(* IEC 61131-3 sources: IRIS-Project/LASAL CONTROL SOFTWARE/LasalProject_2025_09_12/Network/Comunicazione_ModBus, 1 file *)

(* ---- ONE_Comunicazione_ModBus_Table.st ---- *)
#define OBJECTS_CONFIG

//Define part of class _TCPIP_SERVER
#ifndef OS_VERSION_MIN_SALAMANDER
    #define OS_VERSION_MIN_SALAMANDER          0x9000
  #endif
  #define TCP_SVR_NO_ERROR                          0

  #define TCP_SVR_ERR_INVALID_SOCKET            -1

  #define TCP_SVR_ERR_SET_PARA_INVALID_CMD     -10
  #define TCP_SVR_ERR_SET_PARA_INVALID_SUB_CMD -11

  #define TCP_SVR_ERR_TASK_ALREADY_EXIST       -12

  // - RETURN VALUES PRIVATE METHOD Read_AP_TaskPeriod
  #define TCP_SVR_ERR_TASK_TIME_NO_APP            -31
  #define TCP_SVR_ERR_TASK_TIME_WRONG_TASK_TYPE   -33
  #define TCP_SVR_ERR_TASK_TIME_OBJ_NOT_FOUND     -35

  // - RETURN VALUES PRIVATE METHOD Read_LSLOBJ_CRC32
  #define TCP_SVR_ERR_GET_LSLOBJ_NAME             -20
  #define TCP_SVR_ERR_INVALID_POINTER             -21

  // - RETURN VALUES PRIVATE METHOD AP_TaskCreate
  #define TCP_SVR_ERR_TASK_CREATE                 -40

  // - RETURN VALUES PRIVATE METHOD AP_SemaCreate
  #define TCP_SVR_ERR_SEMA_CREATE                 -50
  #define TCP_SVR_ERR_SEMA_INVALID_IDX            -51
  #define TCP_SVR_ERR_SEMA_INVALID_NAME           -52

  #define TCP_SVR_SEND_BUFFER_EMPTY               -6
  #define TCP_SVR_ERR_SEND_BUFFER_FATAL_ERROR     -7

  #define TCP_SVR_SEND_BUFFER_FULL      -4

  #define TCP_SVR_SOCK_INFO_CONNECT                 1
  #define TCP_SVR_SOCK_INFO_DISCONNECT              0

  #define TCP_SVR_ERR_GROUP_OS                      0
  #define TCP_SVR_ERR_GROUP_AP                      1

  #define TCP_SVR_ERR_CODE_AP_TIMEOUT              -1

  #ifndef INIT_FIRSTSCAN
    #define INIT_FIRSTSCAN                         12
  #endif

  #ifndef AP_TASK_PRIORITY_DEFAULT
    #define AP_TASK_PRIORITY_DEFAULT               14
  #endif

  #define TCP_SVR_ERR_MAIN_INIT                   -90

  #define TCP_SVR_ERR_MAX_CONN                    -80

  #ifndef KEEPALIVE_INTERVAL_DEFAULT
    #define KEEPALIVE_INTERVAL_DEFAULT           7200
  #endif

  #ifndef KEEPALIVE_RETRYTIME_DEFAULT
    #define KEEPALIVE_RETRYTIME_DEFAULT            75
  #endif

  #ifndef KEEPALIVE_RETRYCNT_DEFUALT
    #define KEEPALIVE_RETRYCNT_DEFUALT             10
  #endif

  #ifndef CLOSE_SOCKET_TYPE_DEFAULT
    #define CLOSE_SOCKET_TYPE_DEFAULT               0
  #endif
#include "..\..\Class\_TCPIP_SERVER\SalamanderDelay.h"
#include "..\..\Source\MB_Definitions.h"
#include "..\..\Runtime\%LASALAPPDATA%\Runtime\Include\LSL\lsl_st_mt.h"

FUNCTION GLOBAL TAB ONE_Comunicazione_ModBus
-1$UINT, 0$UINT,
0$UINT, 0$UINT,

15$UDINT,
TO_UDINT(916194998), "_CheckSum", 1$UINT, 0$UINT, 3$UINT,
TO_UDINT(1436589033), "_ModBusTCPSLAVE", 1$UINT, 36$UINT, 3$UINT,
TO_UDINT(26234884), "_TCPIP_SERVER", 1$UINT, 38$UINT, 0$UINT,
TO_UDINT(2897291062), "ASCII_BIN", 1$UINT, 21$UINT, 3$UINT,
TO_UDINT(1067997253), "ControlloServerModBus", 0$UINT, 0$UINT, 3$UINT,
TO_UDINT(3132304963), "HoldingRegister", 0$UINT, 0$UINT, 1$UINT,
TO_UDINT(3014633822), "HoldingRegister_2", 0$UINT, 0$UINT, 1$UINT,
TO_UDINT(3299383752), "HoldingRegister_3", 0$UINT, 0$UINT, 1$UINT,
TO_UDINT(418069068), "InputRegister", 0$UINT, 0$UINT, 3$UINT,
TO_UDINT(2225119864), "MerkerEx", 1$UINT, 22$UINT, 9$UINT,
TO_UDINT(3487210139), "MPS", 0$UINT, 0$UINT, 1$UINT,
TO_UDINT(4105514139), "Rack12V", 0$UINT, 0$UINT, 1$UINT,
TO_UDINT(1850111279), "String", 1$UINT, 11$UINT, 9$UINT,
TO_UDINT(2898603620), "StringInternal", 1$UINT, 85$UINT, 0$UINT,
TO_UDINT(3232495061), "VirtualBaseInit", 1$UINT, 3$UINT, 0$UINT,

1$UINT, TO_UDINT(966565638), "_MODBUSTCPSLAVE1\_BASE\CHECKSUM",
1$UINT, TO_UDINT(273951732), "_MODBUSTCPSLAVE2\_BASE\CHECKSUM",
1$UINT, TO_UDINT(3191650917), "_MODBUSTCPSLAVE3\_BASE\CHECKSUM",

_NO_ATTR, TO_UDINT(1516180976), "_MODBUSTCPSLAVE1",
_NO_ATTR, TO_UDINT(3277210698), "_MODBUSTCPSLAVE2",
_NO_ATTR, TO_UDINT(3025237212), "_MODBUSTCPSLAVE3",

_NO_ATTR, TO_UDINT(3586366131), "ASCII_BIN2",
_NO_ATTR, TO_UDINT(2730797605), "ASCII_BIN3",
_NO_ATTR, TO_UDINT(1017134982), "ASCII_BIN4",

_NO_ATTR, TO_UDINT(2237002480), "CONTROLLOSERVERMODBUS1",
_NO_ATTR, TO_UDINT(475833162), "CONTROLLOSERVERMODBUS2",
_NO_ATTR, TO_UDINT(1801163740), "CONTROLLOSERVERMODBUS3",

_NO_ATTR, TO_UDINT(1823689907), "HOLDINGREGISTER1",

_NO_ATTR, TO_UDINT(263994605), "HOLDINGREGISTER_21",

_NO_ATTR, TO_UDINT(380046764), "HOLDINGREGISTER_31",

_NO_ATTR, TO_UDINT(4239264054), "INPUTREGISTER1",
_NO_ATTR, TO_UDINT(1705465996), "INPUTREGISTER2",
_NO_ATTR, TO_UDINT(312502298), "INPUTREGISTER3",

1$UINT, TO_UDINT(392675759), "_MODBUSTCPSLAVE1\_BASE\STRSEMANAME01\MERKEREX0",
1$UINT, TO_UDINT(2391123886), "_MODBUSTCPSLAVE1\_BASE\STRSEMANAME02\MERKEREX0",
1$UINT, TO_UDINT(2044784268), "_MODBUSTCPSLAVE1\_BASE\STRTASKNAME\MERKEREX0",
1$UINT, TO_UDINT(72349916), "_MODBUSTCPSLAVE2\_BASE\STRSEMANAME01\MERKEREX0",
1$UINT, TO_UDINT(2645401309), "_MODBUSTCPSLAVE2\_BASE\STRSEMANAME02\MERKEREX0",
1$UINT, TO_UDINT(3706226144), "_MODBUSTCPSLAVE2\_BASE\STRTASKNAME\MERKEREX0",
1$UINT, TO_UDINT(178786317), "_MODBUSTCPSLAVE3\_BASE\STRSEMANAME01\MERKEREX0",
1$UINT, TO_UDINT(2471130636), "_MODBUSTCPSLAVE3\_BASE\STRSEMANAME02\MERKEREX0",
1$UINT, TO_UDINT(3220135108), "_MODBUSTCPSLAVE3\_BASE\STRTASKNAME\MERKEREX0",

_NO_ATTR, TO_UDINT(3838738401), "MPS1",

_NO_ATTR, TO_UDINT(3841265751), "RACK12V1",

1$UINT, TO_UDINT(191419237), "_MODBUSTCPSLAVE1\_BASE\STRSEMANAME01",
1$UINT, TO_UDINT(2455864031), "_MODBUSTCPSLAVE1\_BASE\STRSEMANAME02",
1$UINT, TO_UDINT(2184963303), "_MODBUSTCPSLAVE1\_BASE\STRTASKNAME",
1$UINT, TO_UDINT(1886802310), "_MODBUSTCPSLAVE2\_BASE\STRSEMANAME01",
1$UINT, TO_UDINT(3917414460), "_MODBUSTCPSLAVE2\_BASE\STRSEMANAME02",
1$UINT, TO_UDINT(560816718), "_MODBUSTCPSLAVE2\_BASE\STRTASKNAME",
1$UINT, TO_UDINT(4021080600), "_MODBUSTCPSLAVE3\_BASE\STRSEMANAME01",
1$UINT, TO_UDINT(1990558626), "_MODBUSTCPSLAVE3\_BASE\STRSEMANAME02",
1$UINT, TO_UDINT(4136624662), "_MODBUSTCPSLAVE3\_BASE\STRTASKNAME",

//Internal connections
0$UDINT,
21$UDINT,
TO_UDINT(3), "CheckSum", TO_UDINT(0),
TO_UDINT(3), "StrTaskName", TO_UDINT(31),
TO_UDINT(3), "StrSemaName01", TO_UDINT(29),
TO_UDINT(3), "StrSemaName02", TO_UDINT(30),
TO_UDINT(4), "CheckSum", TO_UDINT(1),
TO_UDINT(4), "StrTaskName", TO_UDINT(34),
TO_UDINT(4), "StrSemaName01", TO_UDINT(32),
TO_UDINT(4), "StrSemaName02", TO_UDINT(33),
TO_UDINT(5), "CheckSum", TO_UDINT(2),
TO_UDINT(5), "StrTaskName", TO_UDINT(37),
TO_UDINT(5), "StrSemaName01", TO_UDINT(35),
TO_UDINT(5), "StrSemaName02", TO_UDINT(36),
TO_UDINT(29), "MerkerEx0", TO_UDINT(18),
TO_UDINT(30), "MerkerEx0", TO_UDINT(19),
TO_UDINT(31), "MerkerEx0", TO_UDINT(20),
TO_UDINT(32), "MerkerEx0", TO_UDINT(21),
TO_UDINT(33), "MerkerEx0", TO_UDINT(22),
TO_UDINT(34), "MerkerEx0", TO_UDINT(23),
TO_UDINT(35), "MerkerEx0", TO_UDINT(24),
TO_UDINT(36), "MerkerEx0", TO_UDINT(25),
TO_UDINT(37), "MerkerEx0", TO_UDINT(26),
0$UDINT,
21$UDINT,
TO_UDINT(3), "cTable", TO_UDINT(12), "ClassSvr",
TO_UDINT(3), "cTableInputReg", TO_UDINT(15), "ClassSvr",
TO_UDINT(3), "to_AsciiBin", TO_UDINT(6), "Obj_channel",
TO_UDINT(4), "cTable", TO_UDINT(13), "ClassSvr",
TO_UDINT(4), "cTableInputReg", TO_UDINT(16), "ClassSvr",
TO_UDINT(4), "to_AsciiBin", TO_UDINT(7), "Obj_channel",
TO_UDINT(5), "cTable", TO_UDINT(14), "ClassSvr",
TO_UDINT(5), "cTableInputReg", TO_UDINT(17), "ClassSvr",
TO_UDINT(5), "to_AsciiBin", TO_UDINT(8), "Obj_channel",
TO_UDINT(9), "oc_ModBusTCPSlave", TO_UDINT(3), "sControl",
TO_UDINT(10), "oc_ModBusTCPSlave", TO_UDINT(4), "sControl",
TO_UDINT(11), "oc_ModBusTCPSlave", TO_UDINT(5), "sControl",
TO_UDINT(29), "DataBuffer", TO_UDINT(18), "m_udLength",
TO_UDINT(30), "DataBuffer", TO_UDINT(19), "m_udLength",
TO_UDINT(31), "DataBuffer", TO_UDINT(20), "m_udLength",
TO_UDINT(32), "DataBuffer", TO_UDINT(21), "m_udLength",
TO_UDINT(33), "DataBuffer", TO_UDINT(22), "m_udLength",
TO_UDINT(34), "DataBuffer", TO_UDINT(23), "m_udLength",
TO_UDINT(35), "DataBuffer", TO_UDINT(24), "m_udLength",
TO_UDINT(36), "DataBuffer", TO_UDINT(25), "m_udLength",
TO_UDINT(37), "DataBuffer", TO_UDINT(26), "m_udLength",

//Initialization values
0$UDINT,
39$UDINT,
TO_UDINT(3), "sDisable", TO_UDINT(0),//|Comunicazione_ModBus._ModBusTCPSLAVE1.sDisable;
TO_UDINT(3), "cPort", TO_UDINT(502),//|Comunicazione_ModBus._ModBusTCPSLAVE1.cPort;
TO_UDINT(3), "cMaxConnections", TO_UDINT(0),//|Comunicazione_ModBus._ModBusTCPSLAVE1.cMaxConnections;
TO_UDINT(3), "cBufSize", TO_UDINT(100),//|Comunicazione_ModBus._ModBusTCPSLAVE1.cBufSize;
TO_UDINT(3), "cBufSizeInputReg", TO_UDINT(100),//|Comunicazione_ModBus._ModBusTCPSLAVE1.cBufSizeInputReg;
TO_UDINT(3), "cFileOrTable", TO_UDINT(2#11),//|Comunicazione_ModBus._ModBusTCPSLAVE1.cFileOrTable;
TO_UDINT(3), "cTurnBytes", TO_UDINT(1),//|Comunicazione_ModBus._ModBusTCPSLAVE1.cTurnBytes;
TO_UDINT(4), "sDisable", TO_UDINT(0),//|Comunicazione_ModBus._ModBusTCPSLAVE2.sDisable;
TO_UDINT(4), "cPort", TO_UDINT(503),//|Comunicazione_ModBus._ModBusTCPSLAVE2.cPort;
TO_UDINT(4), "cMaxConnections", TO_UDINT(0),//|Comunicazione_ModBus._ModBusTCPSLAVE2.cMaxConnections;
TO_UDINT(4), "cBufSize", TO_UDINT(100),//|Comunicazione_ModBus._ModBusTCPSLAVE2.cBufSize;
TO_UDINT(4), "cBufSizeInputReg", TO_UDINT(100),//|Comunicazione_ModBus._ModBusTCPSLAVE2.cBufSizeInputReg;
TO_UDINT(4), "cFileOrTable", TO_UDINT(2#11),//|Comunicazione_ModBus._ModBusTCPSLAVE2.cFileOrTable;
TO_UDINT(4), "cTurnBytes", TO_UDINT(1),//|Comunicazione_ModBus._ModBusTCPSLAVE2.cTurnBytes;
TO_UDINT(5), "sDisable", TO_UDINT(0),//|Comunicazione_ModBus._ModBusTCPSLAVE3.sDisable;
TO_UDINT(5), "cPort", TO_UDINT(504),//|Comunicazione_ModBus._ModBusTCPSLAVE3.cPort;
TO_UDINT(5), "cMaxConnections", TO_UDINT(0),//|Comunicazione_ModBus._ModBusTCPSLAVE3.cMaxConnections;
TO_UDINT(5), "cBufSize", TO_UDINT(100),//|Comunicazione_ModBus._ModBusTCPSLAVE3.cBufSize;
TO_UDINT(5), "cBufSizeInputReg", TO_UDINT(100),//|Comunicazione_ModBus._ModBusTCPSLAVE3.cBufSizeInputReg;
TO_UDINT(5), "cFileOrTable", TO_UDINT(2#11),//|Comunicazione_ModBus._ModBusTCPSLAVE3.cFileOrTable;
TO_UDINT(5), "cTurnBytes", TO_UDINT(1),//|Comunicazione_ModBus._ModBusTCPSLAVE3.cTurnBytes;
TO_UDINT(18), "ThreadSafe", TO_UDINT(0),//|Comunicazione_ModBus.StrSemaName01\_base\_ModBusTCPSLAVE1\MerkerEx0.ThreadSafe;
TO_UDINT(19), "ThreadSafe", TO_UDINT(0),//|Comunicazione_ModBus.StrSemaName02\_base\_ModBusTCPSLAVE1\MerkerEx0.ThreadSafe;
TO_UDINT(20), "ThreadSafe", TO_UDINT(0),//|Comunicazione_ModBus.StrTaskName\_base\_ModBusTCPSLAVE1\MerkerEx0.ThreadSafe;
TO_UDINT(21), "ThreadSafe", TO_UDINT(0),//|Comunicazione_ModBus.StrSemaName01\_base\_ModBusTCPSLAVE2\MerkerEx0.ThreadSafe;
TO_UDINT(22), "ThreadSafe", TO_UDINT(0),//|Comunicazione_ModBus.StrSemaName02\_base\_ModBusTCPSLAVE2\MerkerEx0.ThreadSafe;
TO_UDINT(23), "ThreadSafe", TO_UDINT(0),//|Comunicazione_ModBus.StrTaskName\_base\_ModBusTCPSLAVE2\MerkerEx0.ThreadSafe;
TO_UDINT(24), "ThreadSafe", TO_UDINT(0),//|Comunicazione_ModBus.StrSemaName01\_base\_ModBusTCPSLAVE3\MerkerEx0.ThreadSafe;
TO_UDINT(25), "ThreadSafe", TO_UDINT(0),//|Comunicazione_ModBus.StrSemaName02\_base\_ModBusTCPSLAVE3\MerkerEx0.ThreadSafe;
TO_UDINT(26), "ThreadSafe", TO_UDINT(0),//|Comunicazione_ModBus.StrTaskName\_base\_ModBusTCPSLAVE3\MerkerEx0.ThreadSafe;
TO_UDINT(29), "SingleRealloc", TO_UDINT(1),//|Comunicazione_ModBus._base\_ModBusTCPSLAVE1\StrSemaName01.SingleRealloc;
TO_UDINT(30), "SingleRealloc", TO_UDINT(1),//|Comunicazione_ModBus._base\_ModBusTCPSLAVE1\StrSemaName02.SingleRealloc;
TO_UDINT(31), "SingleRealloc", TO_UDINT(1),//|Comunicazione_ModBus._base\_ModBusTCPSLAVE1\StrTaskName.SingleRealloc;
TO_UDINT(32), "SingleRealloc", TO_UDINT(1),//|Comunicazione_ModBus._base\_ModBusTCPSLAVE2\StrSemaName01.SingleRealloc;
TO_UDINT(33), "SingleRealloc", TO_UDINT(1),//|Comunicazione_ModBus._base\_ModBusTCPSLAVE2\StrSemaName02.SingleRealloc;
TO_UDINT(34), "SingleRealloc", TO_UDINT(1),//|Comunicazione_ModBus._base\_ModBusTCPSLAVE2\StrTaskName.SingleRealloc;
TO_UDINT(35), "SingleRealloc", TO_UDINT(1),//|Comunicazione_ModBus._base\_ModBusTCPSLAVE3\StrSemaName01.SingleRealloc;
TO_UDINT(36), "SingleRealloc", TO_UDINT(1),//|Comunicazione_ModBus._base\_ModBusTCPSLAVE3\StrSemaName02.SingleRealloc;
TO_UDINT(37), "SingleRealloc", TO_UDINT(1),//|Comunicazione_ModBus._base\_ModBusTCPSLAVE3\StrTaskName.SingleRealloc;

//Symbolic initialization values
0$UDINT,
0$UDINT,

//Initialization of string values
0$UDINT,
0$UDINT,

//Configuration of tasks (RealTime, Cyclic, Background)
0$UDINT,
0$UDINT,

0$UDINT,
3$UDINT,
TO_UDINT(9), (100)$UDINT, 4194303$DINT, 	//CONTROLLOSERVERMODBUS1
TO_UDINT(10), (100)$UDINT, 4194303$DINT, 	//CONTROLLOSERVERMODBUS2
TO_UDINT(11), (100)$UDINT, 4194303$DINT, 	//CONTROLLOSERVERMODBUS3

0$UDINT,
2$UDINT,
TO_UDINT(27), (100)$UDINT, 4194303$DINT, 	//MPS1
TO_UDINT(28), (100)$UDINT, 4194303$DINT, 	//RACK12V1

//External connections
0$UDINT,
5$UDINT,
TO_UDINT(27), "To_Manager_Motori", C_DIR, TO_UDINT(3162257760), "ManagerMotori1","From_MPS",
TO_UDINT(27), "ACKFromMPS", C_DIR, TO_UDINT(2516706254), "DI1601","Input1",
TO_UDINT(27), "c_ReqToMPS", C_DIR, TO_UDINT(1390357230), "TO1271","Output9",
TO_UDINT(27), "To_CameraAlignment_Power", C_DIR, TO_UDINT(2510002277), "ST1516","MaxCurrent",
TO_UDINT(28), "ToPLC", C_DIR, TO_UDINT(1390357230), "TO1271","Output4",

//Magic internal connections
0$UDINT,
0$UDINT,

//Configuration of timeslots of tasks (RealTime, Cyclic)
#ifdef __LSLLDR_TIMESLOTS__
0$UDINT,
0$UDINT,

0$UDINT,
0$UDINT,

#endif //__LSLLDR_TIMESLOTS__

//MultiMaster connections
#ifdef __LSLLDR_MULTIMASTER__
0$UDINT,
0$UDINT,
#endif //__LSLLDR_MULTIMASTER__

//Configuration for task ID (RealTime, CyclicTime)
#ifdef __LSLLDR_TASKID__
"\\\\TASKS2  "
0$UDINT,
0$UDINT,

0$UDINT,
3$UDINT,
(0)$UDINT, 	//CONTROLLOSERVERMODBUS1
(0)$UDINT, 	//CONTROLLOSERVERMODBUS2
(0)$UDINT, 	//CONTROLLOSERVERMODBUS3

0$UDINT,
2$UDINT,
(0)$UDINT, 	//MPS1
(0)$UDINT, 	//RACK12V1

#endif //__LSLLDR_TASKID__

END_FUNCTION
